Fanuc KAREL source: KB00124.KL

PROGRAM KB00124
%NOLOCKGROUP
%ENVIRONMENT FLBT
VAR
  P1: STRING[80]
  P2: INTEGER
BEGIN
  P1 = 'A'
  P2 = 1
  MSG_CONNECT(P1, P2)
END KB00124
